(* IEC 61131-3 sources: rusty/tests/integration/data/empty_proj/src, 2 files *)

(* ---- globals.gvl ---- *)
VAR_GLOBAL
END_VAR

(* ---- mainProg.st ---- *)
PROGRAM mainProg
VAR
x : DINT;
END_VAR

x := 1;
END_PROGRAM
